GLOBALCONSTANTS FileServer (* Konstanten für Übungen 156-159 (File Server) *)
  (* Standard: 61499-1; Description: Copyright (c) 2026 Meisterschulen am Ostbahnhof This program and the accompanying materials are made available under the terms of the Eclipse Public License 2.0 which is available at https://www.eclipse.org/legal/epl-2.0/ SPDX-License-Identifier: EPL-2.0 *)
  (* Version 1.0, 2026-11-25, Franz Höpfinger, Meisterschulen am Ostbahnhof, File Server Filter und Testdateien *)
  PACKAGE Uebungen::const::Uebung_150_159;
  IMPORT isobus::pgn::NAMEFIELD_T;
  VAR_GLOBAL CONSTANT
    FS_ADD : isobus::pgn::NAMEFIELD_T := (bSelfConf := TRUE, bIndGroup := 0, bDevClassInst := 0, bDevClass := 0, bReserved := FALSE, bFunction := 61, bFunctionInst := 0, bEcuInstance := 0, wManufCode := 0, dwIdentNumb := 0); (* File Server: Funktion 61 *)
    FS_FLT : isobus::pgn::NAMEFIELD_T := (bSelfConf := FALSE, bIndGroup := 0, bDevClassInst := 0, bDevClass := 0, bReserved := FALSE, bFunction := 16#FF, bFunctionInst := 0, bEcuInstance := 0, wManufCode := 0, dwIdentNumb := 0); (* prüft nur bFunction *)
    FS_DATEI : STRING := 'logibus_test.txt'; (* Testdatei, relativ zum aktuellen Volume *)
    FS_DATEI_2 : STRING := 'logibus_test2.txt'; (* Kopie zurück auf den File Server *)
    FS_LOKAL : STRING := '/data/fs/logibus_test.txt'; (* lokale Kopie im logiBUS *)
    FS_TEXT : STRING := 'logiBUS File Server Test'; (* Inhalt der Testdatei *)
    FS_WURZEL : STRING := '.'; (* Wurzel des aktuellen Volumes *)
    FS_ORDNER : STRING := 'logibus_test_dir'; (* Testordner Übung 158 *)
    FS_A : STRING := 'logibus_test_dir\a.txt'; (* Übung 158: FsPut-Ziel *)
    FS_B : STRING := 'logibus_test_dir\b.txt'; (* Übung 158: umbenannt *)
    FS_C : STRING := 'logibus_test_dir\c.txt'; (* Übung 158: Kopie *)
    FS_ADD_LOGIBUS : isobus::pgn::NAMEFIELD_T := (bSelfConf := TRUE, bIndGroup := 0, bDevClassInst := 0, bDevClass := 0, bReserved := FALSE, bFunction := 61, bFunctionInst := 0, bEcuInstance := 0, wManufCode := 1116, dwIdentNumb := 0); (* logiBUS-Server, Hersteller 1116 *)
    FS_FLT_LOGIBUS : isobus::pgn::NAMEFIELD_T := (bSelfConf := FALSE, bIndGroup := 0, bDevClassInst := 0, bDevClass := 0, bReserved := FALSE, bFunction := 16#FF, bFunctionInst := 0, bEcuInstance := 0, wManufCode := 16#07FF, dwIdentNumb := 0); (* prüft Funktion und Hersteller *)
    FS_LOGIBUS_ORDNER : STRING := '\\LOGIBUS\IMPORT'; (* Übung 159b: Ordner am logiBUS-Server *)
    FS_LOGIBUS_DATEI : STRING := '\\LOGIBUS\IMPORT\test.txt'; (* Übung 159b: Ziel am logiBUS-Server *)
    FS_LOKAL_ZURUECK : STRING := '/data/fs/logibus_test_zurueck.txt'; (* Übung 159b: zurückgeholte Kopie *)
  END_VAR
END_GLOBALCONSTANTS
